{attribute 'TcGenerated'}
{attribute 'no-analysis'}
{attribute 'linkalways'}
// This function has been automatically generated from the project information.
VAR_GLOBAL CONSTANT
	{attribute 'const_non_replaced'}
	stLibVersion_Intecre_TwinSAFE_Models : ST_LibVersion := (iMajor := 0, iMinor := 5, iBuild := 0, iRevision := 3, nFlags := 0, sVersion := '0.5.0.3');
END_VAR

(* stored: Version 1.1.0.1
   GVL Global_Version: Id {29903f6a-70f9-4ef0-b109-88f6b3657356} *)
